FUNCTION_BLOCK TcoState EXTENDS TcoStateBase

METHOD PUBLIC ChangeState : ITcoState
VAR_INPUT
	NewState : INT;
END_VAR
ChangeState := SUPER^.ChangeStateProtected(NewState);
END_METHOD

(*~
	<docu>
		<summary>
			This method is called on each change of the <c>State</c>. This method could be overloaded and custom code should be placed here.	
		</summary>			
	</docu>	
~*)
METHOD PROTECTED OnStateChange
VAR_INPUT
	PreviousState	: INT;
	NewState 		: INT;
END_VAR
SUPER^.OnStateChange(PreviousState, NewState);
END_METHOD

END_FUNCTION_BLOCK

(* stored: Version 1.1.0.1
   POU TcoState: Id {e15c5fcf-81d3-038e-202e-1cd87b834ace}, SpecialFunc None
   Method ChangeState: Id {8a2449de-98e2-0003-0ff6-3dd7ed17800f}
   Method OnStateChange: Id {3086bfc0-6684-0c18-3a68-e8c47053ddcc} *)
